(* IEC 61131-3 sources: llm-plc-st-eval/data/definitivo/gemini-3.1-pro-preview/C3/zero_shot, 3 files *)

(* ---- ejec_1.st ---- *)
```iecst
PROGRAM PRG_Conversion
VAR_INPUT
    btnMarcha : BOOL; // Botón de inicio (contacto normalmente abierto)
    btnParo : BOOL;   // Botón de detención (contacto normalmente cerrado en la lógica)
END_VAR

VAR_OUTPUT
    motor : BOOL;     // Salida para el motor
    lampara : BOOL;   // Salida para la lámpara indicadora
END_VAR

VAR
    T1 : TON;         // Temporizador de retardo a la conexión
END_VAR

// Rama 1: Lógica de arranque y enclavamiento del motor
motor := (btnMarcha OR motor) AND NOT btnParo;

// Rama 2: Llamada al temporizador TON (10 segundos) activado por el motor
T1(IN := motor, PT := T#10S);

// Rama 3: Activación de la lámpara cuando el temporizador finaliza
lampara := T1.Q;

END_PROGRAM
```

(* ---- ejec_2.st ---- *)
```iecst
PROGRAM PRG_Conversion
VAR_INPUT
    btnMarcha : BOOL; // Contacto normalmente abierto para iniciar
    btnParo : BOOL;   // Contacto normalmente cerrado para detener
END_VAR

VAR_OUTPUT
    motor : BOOL;     // Bobina del motor
    lampara : BOOL;   // Bobina de la lámpara indicadora
END_VAR

VAR
    T1 : TON;         // Temporizador a la conexión (Timer On Delay)
END_VAR

// Rama 1: Lógica de enclavamiento (arranque y paro) para el motor
motor := (btnMarcha OR motor) AND NOT btnParo;

// Rama 2: Llamada al temporizador T1, se activa cuando el motor está encendido
T1(IN := motor, PT := T#10S);

// Rama 3: La lámpara se enciende cuando el temporizador T1 termina su conteo
lampara := T1.Q;

END_PROGRAM
```

(* ---- ejec_3.st ---- *)
```iecst
PROGRAM PRG_Conversion
VAR_INPUT
    btnMarcha : BOOL; // Contacto normalmente abierto para arranque
    btnParo : BOOL;   // Contacto normalmente cerrado para detención
END_VAR

VAR_OUTPUT
    motor : BOOL;     // Bobina del motor
    lampara : BOOL;   // Bobina de la lámpara
END_VAR

VAR
    T1 : TON;         // Temporizador de retardo a la conexión
END_VAR

// Rama 1: Circuito de auto-retención (enclavamiento) del motor
motor := (btnMarcha OR motor) AND NOT btnParo;

// Rama 2: El motor activa el temporizador TON con un preset de 10 segundos
T1(IN := motor, PT := T#10S);

// Rama 3: La salida del temporizador enciende la lámpara
lampara := T1.Q;

END_PROGRAM
```
